SUBAPPLICATION Uebung_094b4_AX (* Wie Uebung_094b_AX, aber mit MyLib_AX::sys::NumericValue_TO_AUI2 als wiederverwendbarem Baustein statt der inline verdrahteten Kette (NumericValue_IDA+AD_TO_AUI+AUI_TO_AUI2+AUI_TO_AUDI+Q_NumericValue_AUDI). *)
  (* Standard: 61499-2; Description: Copyright (c) 2026 Meisterschulen am Ostbahnhof This program and the accompanying materials are made available under the terms of the Eclipse Public License 2.0 which is available at https://www.eclipse.org/legal/epl-2.0/ SPDX-License-Identifier: EPL-2.0 *)
  (* Version 1.0, 2026-10-13, Franz Höpfinger, Meisterschulen am Ostbahnhof, 2. Version von Uebung_094b_AX: die Lese/Echo-Kette wurde nach MyLib_AX::sys::NumericValue_TO_AUI2 ausgelagert (u16ObjId als SubApp-Parameter statt fest verdrahtet), analog Uebung_094b3_AX/Uebung_094c2_AX. *)
  PACKAGE Uebungen;
  IMPORT Uebungen::const::UT::DefaultPool::InputNumber_I1;
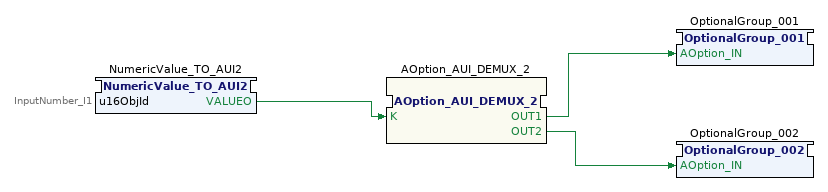
  FBS
    AOption_AUI_DEMUX_2 : Option::selection::AOption_AUI_DEMUX_2;
  END_FBS
  SUBAPPS
    NumericValue_TO_AUI2 : MyLib::sys::NumericValue_TO_AUI2(u16ObjId := InputNumber_I1);
    OptionalGroup_001 : MyLib_AX_Option::sys::OptionalGroup_001;
    OptionalGroup_002 : MyLib_AX_Option::sys::OptionalGroup_002;
  END_SUBAPPS
  ADAPTER_CONNECTIONS
    NumericValue_TO_AUI2.VALUEO TO AOption_AUI_DEMUX_2.K;
    AOption_AUI_DEMUX_2.OUT1 TO OptionalGroup_001.AOption_IN;
    AOption_AUI_DEMUX_2.OUT2 TO OptionalGroup_002.AOption_IN;
  END_CONNECTIONS
END_SUBAPPLICATION
